{attribute 'no_assign'}
FUNCTION_BLOCK FB_DO_WTURBINE_LD0_WYAW1_YwAngSpt EXTENDS FB_AcsiCommonDataClass
VAR_INPUT
	val: FB_DO_WTURBINE_LD0_WYAW1_YwAngSpt_val := (sClass:='APC', bLinkResult:=THIS^.AddDataToContainer(ipData:=val));
END_VAR
VAR
END_VAR

END_FUNCTION_BLOCK

(* stored: Version 1.1.0.1
   POU FB_DO_WTURBINE_LD0_WYAW1_YwAngSpt: Id {2c3704b0-415e-41c7-b252-3f6a8a7e767a}, SpecialFunc None *)
